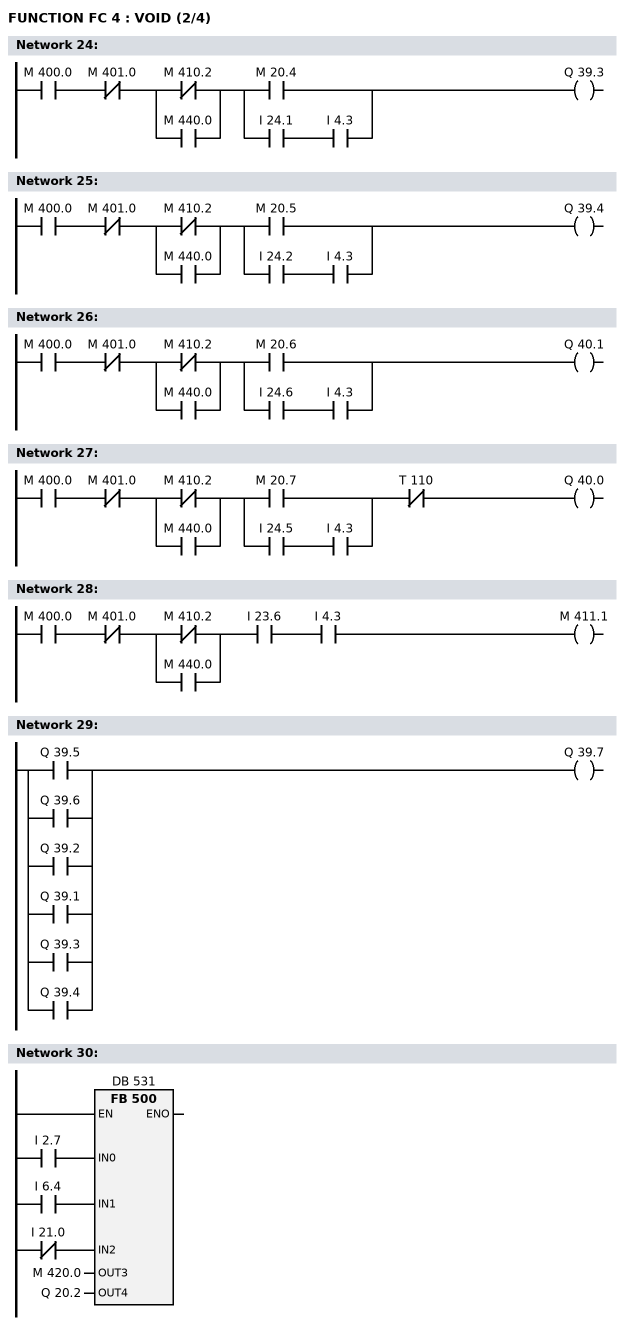

      A     M    400.0;
      AN    M    401.0;
      A(    ;
      ON    M    410.2;
      O     M    440.0;
      )     ;
      A(    ;
      O     M     20.4;
      O     ;
      A     I     24.1;
      A     I      4.3;
      )     ;
      =     Q     39.3;
NETWORK
TITLE =

      A     M    400.0;
      AN    M    401.0;
      A(    ;
      ON    M    410.2;
      O     M    440.0;
      )     ;
      A(    ;
      O     M     20.5;
      O     ;
      A     I     24.2;
      A     I      4.3;
      )     ;
      =     Q     39.4;
NETWORK
TITLE =

      A     M    400.0;
      AN    M    401.0;
      A(    ;
      ON    M    410.2;
      O     M    440.0;
      )     ;
      A(    ;
      O     M     20.6;
      O     ;
      A     I     24.6;
      A     I      4.3;
      )     ;
      =     Q     40.1;
NETWORK
TITLE =

      A     M    400.0;
      AN    M    401.0;
      A(    ;
      ON    M    410.2;
      O     M    440.0;
      )     ;
      A(    ;
      O     M     20.7;
      O     ;
      A     I     24.5;
      A     I      4.3;
      )     ;
      AN    T    110;
      =     Q     40.0;
NETWORK
TITLE =

      A     M    400.0;
      AN    M    401.0;
      A(    ;
      ON    M    410.2;
      O     M    440.0;
      )     ;
      A     I     23.6;
      A     I      4.3;
      =     M    411.1;
NETWORK
TITLE =

      O     Q     39.5;
      O     Q     39.6;
      O     Q     39.2;
      O     Q     39.1;
      O     Q     39.3;
      O     Q     39.4;
      =     Q     39.7;
NETWORK
TITLE =

      A     I      2.7;
      =     L      0.0;
      BLD   103;
      A     I      6.4;
      =     L      0.1;
      BLD   103;
      AN    I     21.0;
      =     L      0.2;
      BLD   103;
      CALL FB   500 , DB   531 (
           IN0                      := L      0.0,
           IN1                      := L      0.1,
           IN2                      := L      0.2,
           OUT3                     := M    420.0,
           OUT4                     := Q     20.2);
      NOP   0;
NETWORK
TITLE =
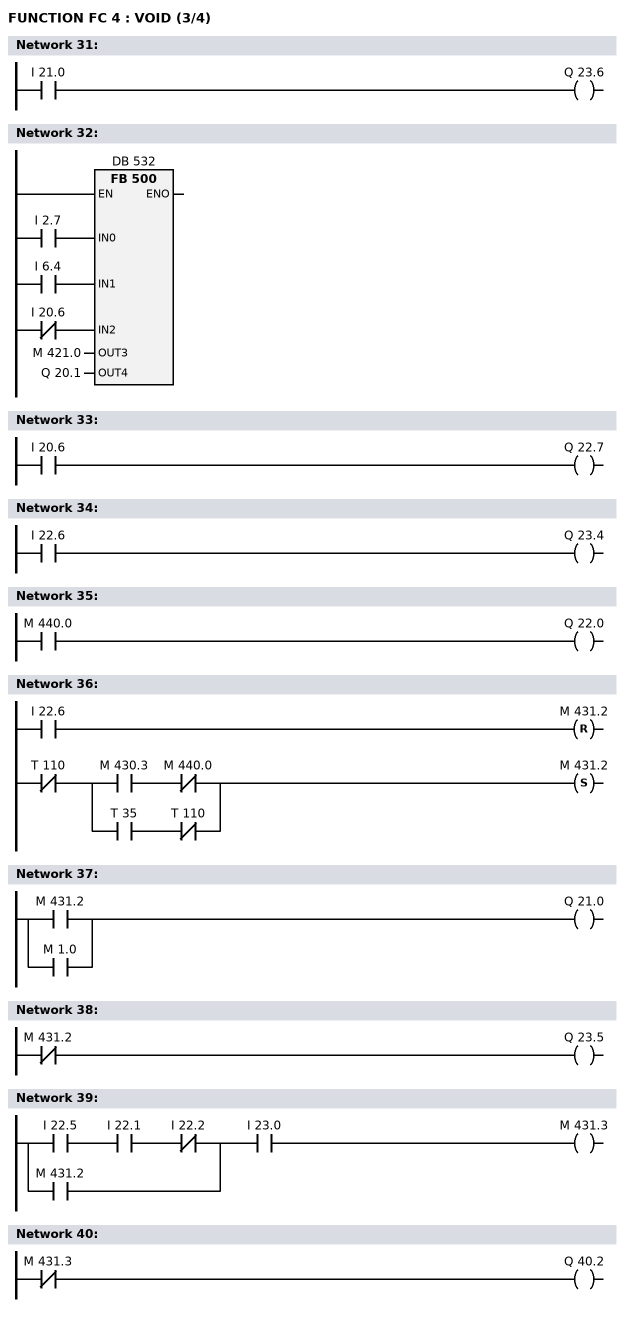

      A     I     21.0;
      =     Q     23.6;
NETWORK
TITLE =

      A     I      2.7;
      =     L      0.0;
      BLD   103;
      A     I      6.4;
      =     L      0.1;
      BLD   103;
      AN    I     20.6;
      =     L      0.2;
      BLD   103;
      CALL FB   500 , DB   532 (
           IN0                      := L      0.0,
           IN1                      := L      0.1,
           IN2                      := L      0.2,
           OUT3                     := M    421.0,
           OUT4                     := Q     20.1);
      NOP   0;
NETWORK
TITLE =

      A     I     20.6;
      =     Q     22.7;
NETWORK
TITLE =

      A     I     22.6;
      =     Q     23.4;
NETWORK
TITLE =

      A     M    440.0;
      =     Q     22.0;
NETWORK
TITLE =

      A     I     22.6;
      R     M    431.2;
      AN    T    110;
      A(    ;
      A     M    430.3;
      AN    M    440.0;
      O     ;
      A     T     35;
      AN    T    110;
      )     ;
      S     M    431.2;
      NOP   0;
NETWORK
TITLE =

      O     M    431.2;
      O     M      1.0;
      =     Q     21.0;
NETWORK
TITLE =

      AN    M    431.2;
      =     Q     23.5;
NETWORK
TITLE =

      A(    ;
      A     I     22.5;
      A     I     22.1;
      AN    I     22.2;
      O     M    431.2;
      )     ;
      A     I     23.0;
      =     M    431.3;
NETWORK
TITLE =

      AN    M    431.3;
      =     Q     40.2;
NETWORK
TITLE =
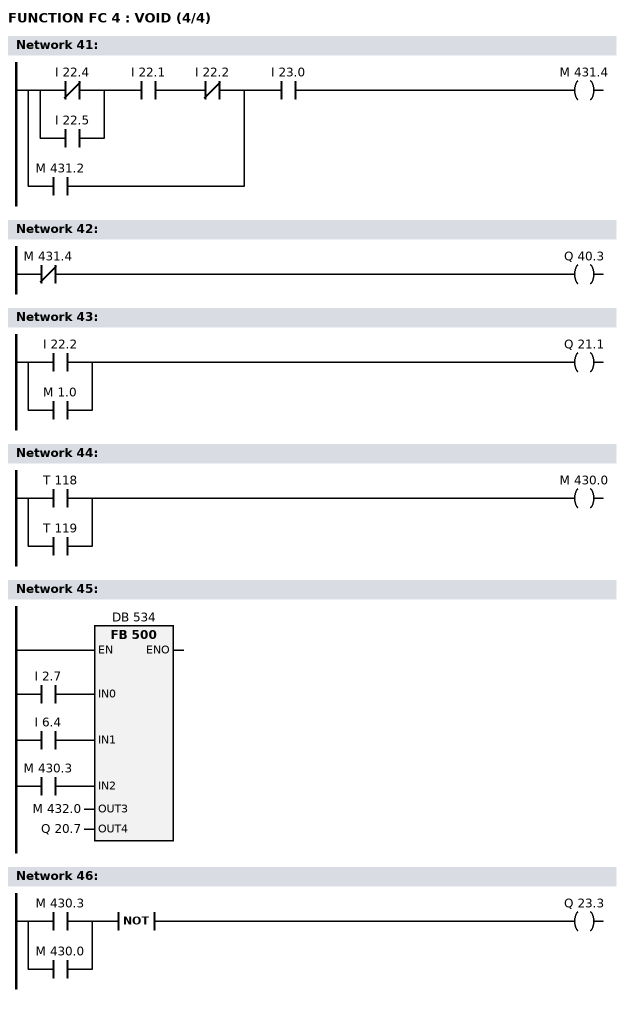

      A(    ;
      A(    ;
      ON    I     22.4;
      O     I     22.5;
      )     ;
      A     I     22.1;
      AN    I     22.2;
      O     M    431.2;
      )     ;
      A     I     23.0;
      =     M    431.4;
NETWORK
TITLE =

      AN    M    431.4;
      =     Q     40.3;
NETWORK
TITLE =

      O     I     22.2;
      O     M      1.0;
      =     Q     21.1;
NETWORK
TITLE =

      O     T    118;
      O     T    119;
      =     M    430.0;
NETWORK
TITLE =

      A     I      2.7;
      =     L      0.0;
      BLD   103;
      A     I      6.4;
      =     L      0.1;
      BLD   103;
      A     M    430.3;
      =     L      0.2;
      BLD   103;
      CALL FB   500 , DB   534 (
           IN0                      := L      0.0,
           IN1                      := L      0.1,
           IN2                      := L      0.2,
           OUT3                     := M    432.0,
           OUT4                     := Q     20.7);
      NOP   0;
NETWORK
TITLE =

      A(    ;
      O     M    430.3;
      O     M    430.0;
      )     ;
      NOT   ;
      =     Q     23.3;
NETWORK
TITLE =

      A(    ;
      A     I     21.5;
      L     S5T#150MS;
      SD    T    103;
      NOP   0;
      NOP   0;
      NOP   0;
      A     T    103;
      )     ;
      NOT   ;
      =     Q     21.6;
NETWORK
TITLE =

      A(    ;
      A     I     21.7;
      L     S5T#150MS;
      SD    T    104;
      NOP   0;
      NOP   0;
      NOP   0;
      A     T    104;
      )     ;
      NOT   ;
      =     Q     23.1;
NETWORK
TITLE =

      A(    ;
      A     I     21.6;
      L     S5T#150MS;
      SD    T    106;
      NOP   0;
      NOP   0;
      NOP   0;
      A     T    106;
      )     ;
      NOT   ;
      =     Q     22.6;
NETWORK
TITLE =

      A(    ;
      A     I     21.4;
      L     S5T#150MS;
      SD    T    107;
      NOP   0;
      NOP   0;
      NOP   0;
      A     T    107;
      )     ;
      NOT   ;
      =     Q     23.2;
NETWORK
TITLE =
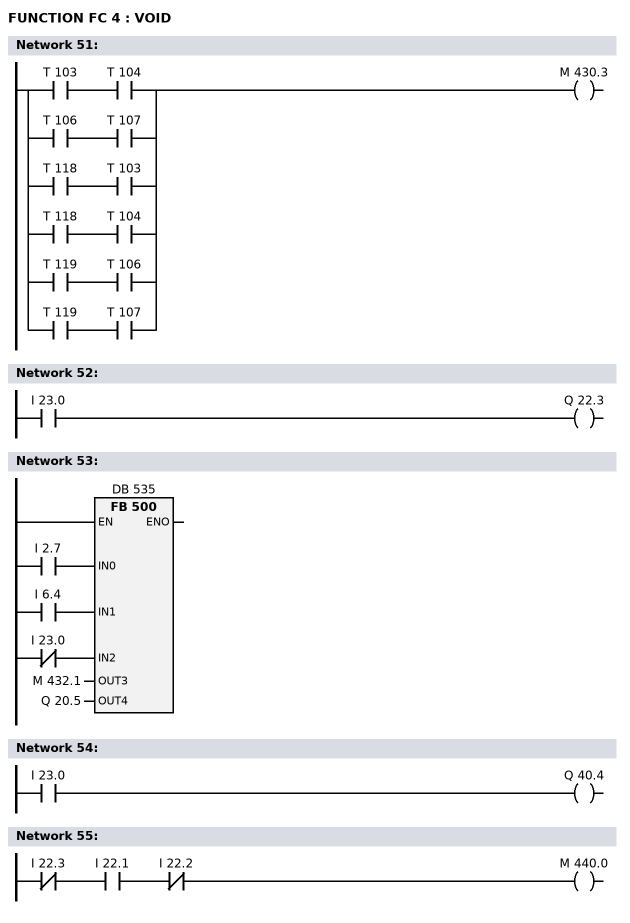

      A     T    103;
      A     T    104;
      O     ;
      A     T    106;
      A     T    107;
      O     ;
      A     T    118;
      A     T    103;
      O     ;
      A     T    118;
      A     T    104;
      O     ;
      A     T    119;
      A     T    106;
      O     ;
      A     T    119;
      A     T    107;
      =     M    430.3;
NETWORK
TITLE =

      A     I     23.0;
      =     Q     22.3;
NETWORK
TITLE =

      A     I      2.7;
      =     L      0.0;
      BLD   103;
      A     I      6.4;
      =     L      0.1;
      BLD   103;
      AN    I     23.0;
      =     L      0.2;
      BLD   103;
      CALL FB   500 , DB   535 (
           IN0                      := L      0.0,
           IN1                      := L      0.1,
           IN2                      := L      0.2,
           OUT3                     := M    432.1,
           OUT4                     := Q     20.5);
      NOP   0;
NETWORK
TITLE =

      A     I     23.0;
      =     Q     40.4;
NETWORK
TITLE =

      AN    I     22.3;
      A     I     22.1;
      AN    I     22.2;
      =     M    440.0;
END_FUNCTION

FUNCTION FC 5 : VOID
VERSION : 0.1

BEGIN
NETWORK
TITLE =
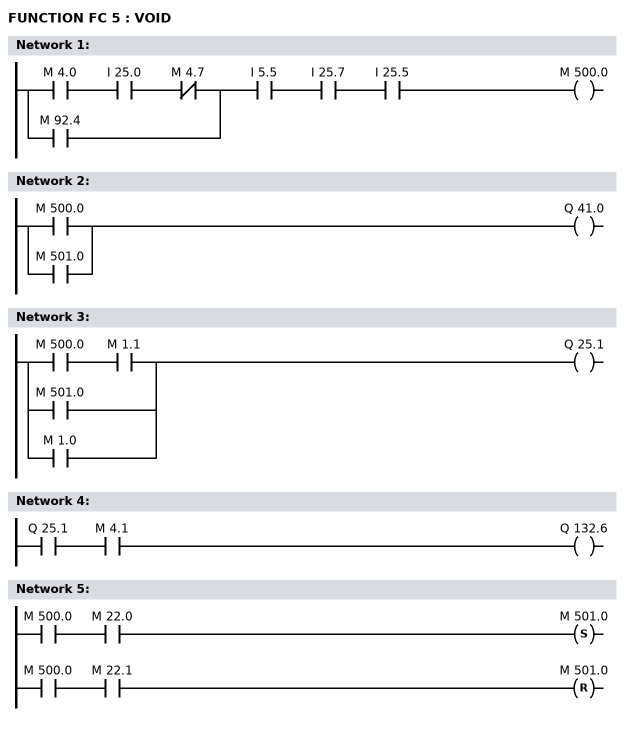

      A(    ;
      A     M      4.0;
      A     I     25.0;
      AN    M      4.7;
      O     M     92.4;
      )     ;
      A     I      5.5;
      A     I     25.7;
      A     I     25.5;
      =     M    500.0;
NETWORK
TITLE =

      O     M    500.0;
      O     M    501.0;
      =     Q     41.0;
NETWORK
TITLE =

      A     M    500.0;
      A     M      1.1;
      O     M    501.0;
      O     M      1.0;
      =     Q     25.1;
NETWORK
TITLE =

      A     Q     25.1;
      A     M      4.1;
      =     Q    132.6;
NETWORK
TITLE =

      A     M    500.0;
      A     M     22.0;
      S     M    501.0;
      A     M    500.0;
      A     M     22.1;
      R     M    501.0;
      NOP   0;
NETWORK
TITLE =

      A(    ;
      A     I     25.3;
      L     S5T#150MS;
      SD    T    128;
      NOP   0;
      NOP   0;
      NOP   0;
      A     T    128;
      )     ;
      NOT   ;
      =     Q     25.7;
NETWORK
TITLE =

      A(    ;
      A     I     25.2;
      L     S5T#150MS;
      SD    T    129;
      NOP   0;
      NOP   0;
      NOP   0;
      A     T    129;
      )     ;
      NOT   ;
      =     Q     25.6;
NETWORK
TITLE =
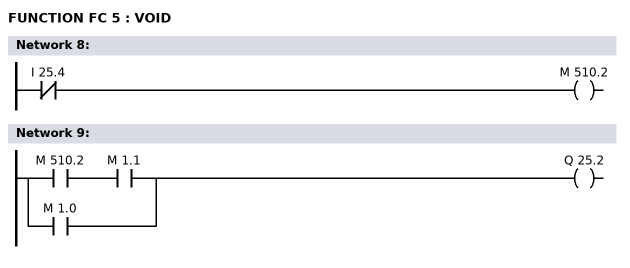

      AN    I     25.4;
      =     M    510.2;
NETWORK
TITLE =

      A     M    510.2;
      A     M      1.1;
      O     M      1.0;
      =     Q     25.2;
NETWORK
TITLE =

      O(    ;
      A     I     25.1;
      L     S5T#150MS;
      SD    T    130;
      NOP   0;
      NOP   0;
      NOP   0;
      A     T    130;
      )     ;
      O     M      1.0;
      =     Q     25.0;
NETWORK
TITLE =
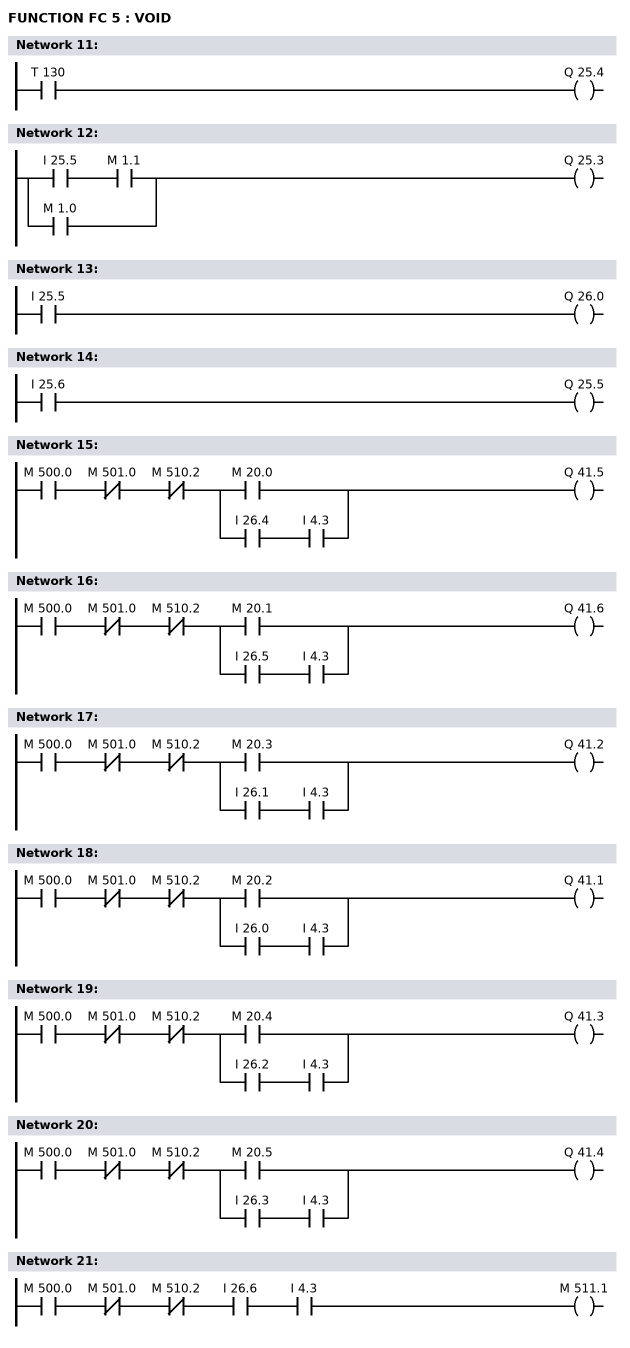

      A     T    130;
      =     Q     25.4;
NETWORK
TITLE =

      A     I     25.5;
      A     M      1.1;
      O     M      1.0;
      =     Q     25.3;
NETWORK
TITLE =

      A     I     25.5;
      =     Q     26.0;
NETWORK
TITLE =

      A     I     25.6;
      =     Q     25.5;
NETWORK
TITLE =

      A     M    500.0;
      AN    M    501.0;
      AN    M    510.2;
      A(    ;
      O     M     20.0;
      O     ;
      A     I     26.4;
      A     I      4.3;
      )     ;
      =     Q     41.5;
NETWORK
TITLE =

      A     M    500.0;
      AN    M    501.0;
      AN    M    510.2;
      A(    ;
      O     M     20.1;
      O     ;
      A     I     26.5;
      A     I      4.3;
      )     ;
      =     Q     41.6;
NETWORK
TITLE =

      A     M    500.0;
      AN    M    501.0;
      AN    M    510.2;
      A(    ;
      O     M     20.3;
      O     ;
      A     I     26.1;
      A     I      4.3;
      )     ;
      =     Q     41.2;
NETWORK
TITLE =

      A     M    500.0;
      AN    M    501.0;
      AN    M    510.2;
      A(    ;
      O     M     20.2;
      O     ;
      A     I     26.0;
      A     I      4.3;
      )     ;
      =     Q     41.1;
NETWORK
TITLE =

      A     M    500.0;
      AN    M    501.0;
      AN    M    510.2;
      A(    ;
      O     M     20.4;
      O     ;
      A     I     26.2;
      A     I      4.3;
      )     ;
      =     Q     41.3;
NETWORK
TITLE =

      A     M    500.0;
      AN    M    501.0;
      AN    M    510.2;
      A(    ;
      O     M     20.5;
      O     ;
      A     I     26.3;
      A     I      4.3;
      )     ;
      =     Q     41.4;
NETWORK
TITLE =

      A     M    500.0;
      AN    M    501.0;
      AN    M    510.2;
      A     I     26.6;
      A     I      4.3;
      =     M    511.1;
END_FUNCTION

FUNCTION FC 6 : VOID
VERSION : 0.1

BEGIN
NETWORK
TITLE =
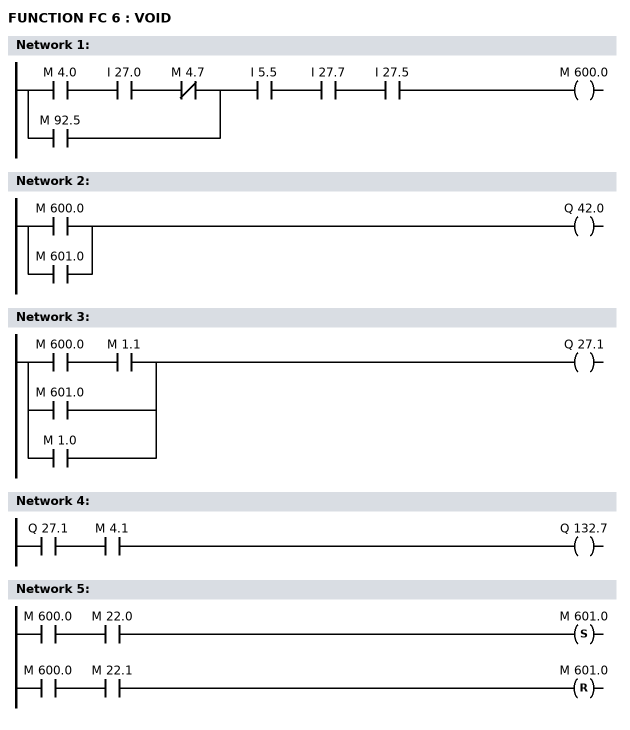

      A(    ;
      A     M      4.0;
      A     I     27.0;
      AN    M      4.7;
      O     M     92.5;
      )     ;
      A     I      5.5;
      A     I     27.7;
      A     I     27.5;
      =     M    600.0;
NETWORK
TITLE =

      O     M    600.0;
      O     M    601.0;
      =     Q     42.0;
NETWORK
TITLE =

      A     M    600.0;
      A     M      1.1;
      O     M    601.0;
      O     M      1.0;
      =     Q     27.1;
NETWORK
TITLE =

      A     Q     27.1;
      A     M      4.1;
      =     Q    132.7;
NETWORK
TITLE =

      A     M    600.0;
      A     M     22.0;
      S     M    601.0;
      A     M    600.0;
      A     M     22.1;
      R     M    601.0;
      NOP   0;
NETWORK
TITLE =

      A(    ;
      A     I     27.3;
      L     S5T#150MS;
      SD    T    148;
      NOP   0;
      NOP   0;
      NOP   0;
      A     T    148;
      )     ;
      NOT   ;
      =     Q     27.7;
NETWORK
TITLE =

      A(    ;
      A     I     27.2;
      L     S5T#150MS;
      SD    T    149;
      NOP   0;
      NOP   0;
      NOP   0;
      A     T    149;
      )     ;
      NOT   ;
      =     Q     27.6;
NETWORK
TITLE =
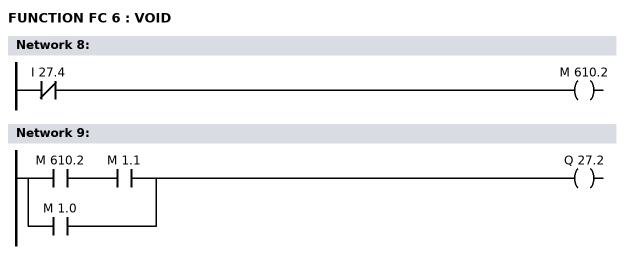

      AN    I     27.4;
      =     M    610.2;
NETWORK
TITLE =

      A     M    610.2;
      A     M      1.1;
      O     M      1.0;
      =     Q     27.2;
NETWORK
TITLE =

      O(    ;
      A     I     27.1;
      L     S5T#150MS;
      SD    T    150;
      NOP   0;
      NOP   0;
      NOP   0;
      A     T    150;
      )     ;
      O     M      1.0;
      =     Q     27.0;
NETWORK
TITLE =
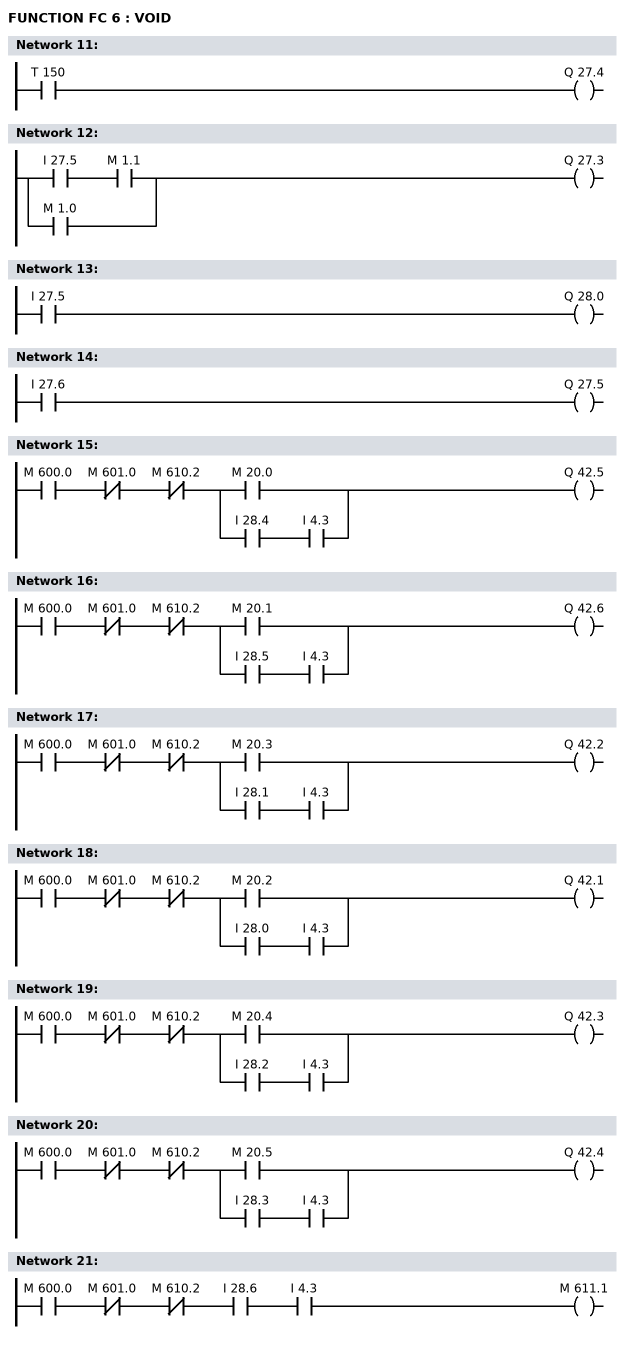

      A     T    150;
      =     Q     27.4;
NETWORK
TITLE =

      A     I     27.5;
      A     M      1.1;
      O     M      1.0;
      =     Q     27.3;
NETWORK
TITLE =

      A     I     27.5;
      =     Q     28.0;
NETWORK
TITLE =

      A     I     27.6;
      =     Q     27.5;
NETWORK
TITLE =

      A     M    600.0;
      AN    M    601.0;
      AN    M    610.2;
      A(    ;
      O     M     20.0;
      O     ;
      A     I     28.4;
      A     I      4.3;
      )     ;
      =     Q     42.5;
NETWORK
TITLE =

      A     M    600.0;
      AN    M    601.0;
      AN    M    610.2;
      A(    ;
      O     M     20.1;
      O     ;
      A     I     28.5;
      A     I      4.3;
      )     ;
      =     Q     42.6;
NETWORK
TITLE =

      A     M    600.0;
      AN    M    601.0;
      AN    M    610.2;
      A(    ;
      O     M     20.3;
      O     ;
      A     I     28.1;
      A     I      4.3;
      )     ;
      =     Q     42.2;
NETWORK
TITLE =

      A     M    600.0;
      AN    M    601.0;
      AN    M    610.2;
      A(    ;
      O     M     20.2;
      O     ;
      A     I     28.0;
      A     I      4.3;
      )     ;
      =     Q     42.1;
NETWORK
TITLE =

      A     M    600.0;
      AN    M    601.0;
      AN    M    610.2;
      A(    ;
      O     M     20.4;
      O     ;
      A     I     28.2;
      A     I      4.3;
      )     ;
      =     Q     42.3;
NETWORK
TITLE =

      A     M    600.0;
      AN    M    601.0;
      AN    M    610.2;
      A(    ;
      O     M     20.5;
      O     ;
      A     I     28.3;
      A     I      4.3;
      )     ;
      =     Q     42.4;
NETWORK
TITLE =

      A     M    600.0;
      AN    M    601.0;
      AN    M    610.2;
      A     I     28.6;
      A     I      4.3;
      =     M    611.1;
END_FUNCTION

FUNCTION FC 7 : VOID
VERSION : 0.1

BEGIN
NETWORK
TITLE =
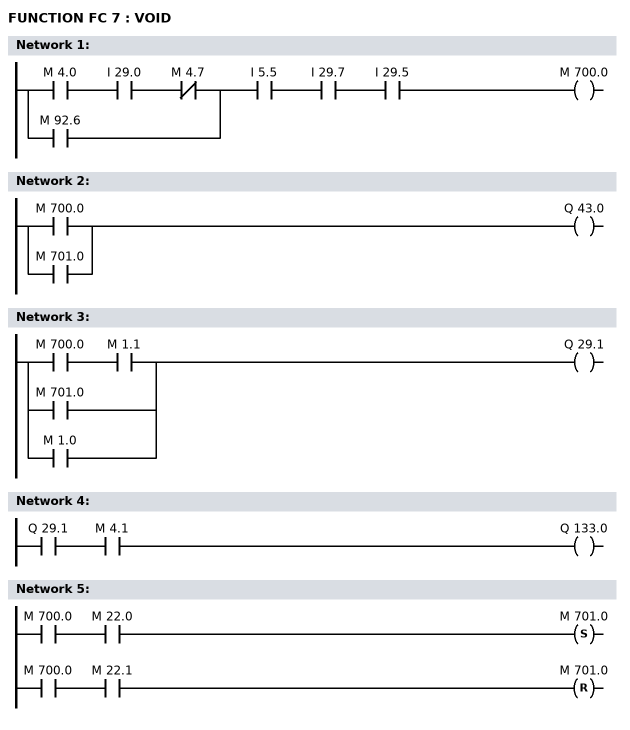

      A(    ;
      A     M      4.0;
      A     I     29.0;
      AN    M      4.7;
      O     M     92.6;
      )     ;
      A     I      5.5;
      A     I     29.7;
      A     I     29.5;
      =     M    700.0;
NETWORK
TITLE =

      O     M    700.0;
      O     M    701.0;
      =     Q     43.0;
NETWORK
TITLE =

      A     M    700.0;
      A     M      1.1;
      O     M    701.0;
      O     M      1.0;
      =     Q     29.1;
NETWORK
TITLE =

      A     Q     29.1;
      A     M      4.1;
      =     Q    133.0;
NETWORK
TITLE =

      A     M    700.0;
      A     M     22.0;
      S     M    701.0;
      A     M    700.0;
      A     M     22.1;
      R     M    701.0;
      NOP   0;
NETWORK
TITLE =

      A(    ;
      A     I     29.3;
      L     S5T#150MS;
      SD    T    168;
      NOP   0;
      NOP   0;
      NOP   0;
      A     T    168;
      )     ;
      NOT   ;
      =     Q     29.7;
NETWORK
TITLE =

      A(    ;
      A     I     29.2;
      L     S5T#150MS;
      SD    T    169;
      NOP   0;
      NOP   0;
      NOP   0;
      A     T    169;
      )     ;
      NOT   ;
      =     Q     29.6;
NETWORK
TITLE =
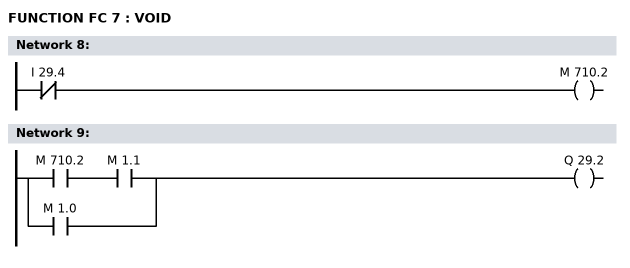

      AN    I     29.4;
      =     M    710.2;
NETWORK
TITLE =

      A     M    710.2;
      A     M      1.1;
      O     M      1.0;
      =     Q     29.2;
NETWORK
TITLE =

      O(    ;
      A     I     29.1;
      L     S5T#150MS;
      SD    T    170;
      NOP   0;
      NOP   0;
      NOP   0;
      A     T    170;
      )     ;
      O     M      1.0;
      =     Q     29.0;
NETWORK
TITLE =
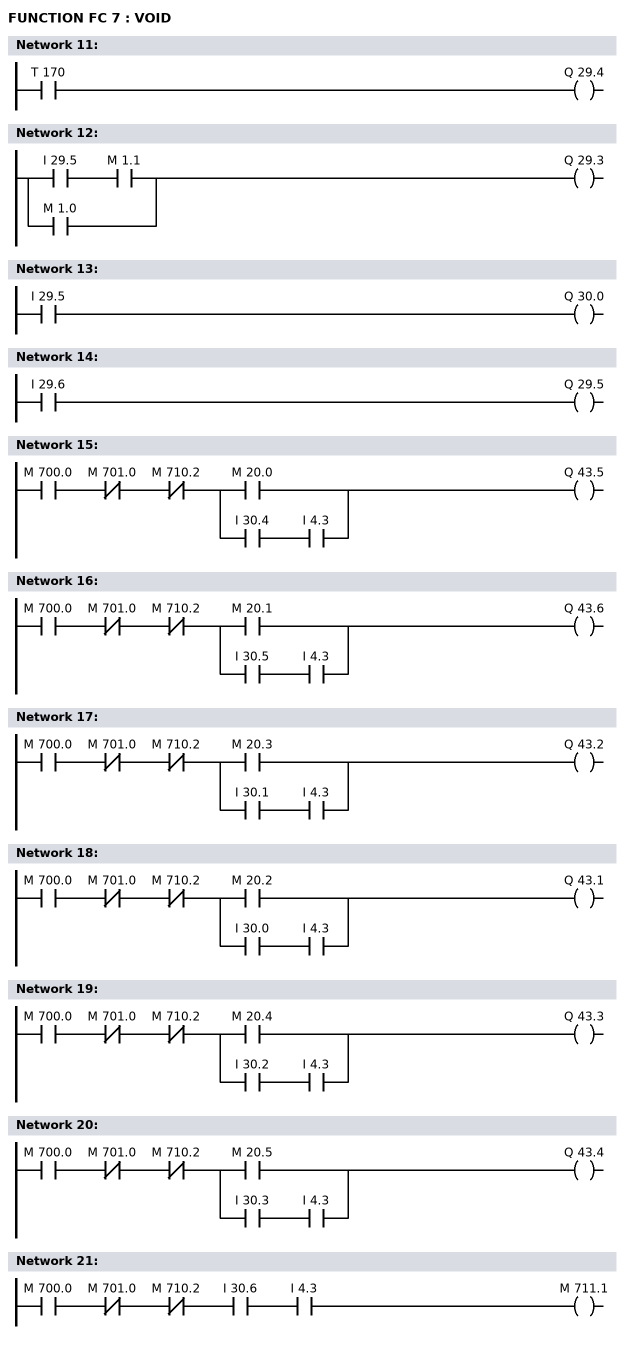

      A     T    170;
      =     Q     29.4;
NETWORK
TITLE =

      A     I     29.5;
      A     M      1.1;
      O     M      1.0;
      =     Q     29.3;
NETWORK
TITLE =

      A     I     29.5;
      =     Q     30.0;
NETWORK
TITLE =

      A     I     29.6;
      =     Q     29.5;
NETWORK
TITLE =

      A     M    700.0;
      AN    M    701.0;
      AN    M    710.2;
      A(    ;
      O     M     20.0;
      O     ;
      A     I     30.4;
      A     I      4.3;
      )     ;
      =     Q     43.5;
NETWORK
TITLE =

      A     M    700.0;
      AN    M    701.0;
      AN    M    710.2;
      A(    ;
      O     M     20.1;
      O     ;
      A     I     30.5;
      A     I      4.3;
      )     ;
      =     Q     43.6;
NETWORK
TITLE =

      A     M    700.0;
      AN    M    701.0;
      AN    M    710.2;
      A(    ;
      O     M     20.3;
      O     ;
      A     I     30.1;
      A     I      4.3;
      )     ;
      =     Q     43.2;
NETWORK
TITLE =

      A     M    700.0;
      AN    M    701.0;
      AN    M    710.2;
      A(    ;
      O     M     20.2;
      O     ;
      A     I     30.0;
      A     I      4.3;
      )     ;
      =     Q     43.1;
NETWORK
TITLE =

      A     M    700.0;
      AN    M    701.0;
      AN    M    710.2;
      A(    ;
      O     M     20.4;
      O     ;
      A     I     30.2;
      A     I      4.3;
      )     ;
      =     Q     43.3;
NETWORK
TITLE =

      A     M    700.0;
      AN    M    701.0;
      AN    M    710.2;
      A(    ;
      O     M     20.5;
      O     ;
      A     I     30.3;
      A     I      4.3;
      )     ;
      =     Q     43.4;
NETWORK
TITLE =

      A     M    700.0;
      AN    M    701.0;
      AN    M    710.2;
      A     I     30.6;
      A     I      4.3;
      =     M    711.1;
END_FUNCTION

FUNCTION FC 11 : VOID
VERSION : 0.1

BEGIN
NETWORK
TITLE =
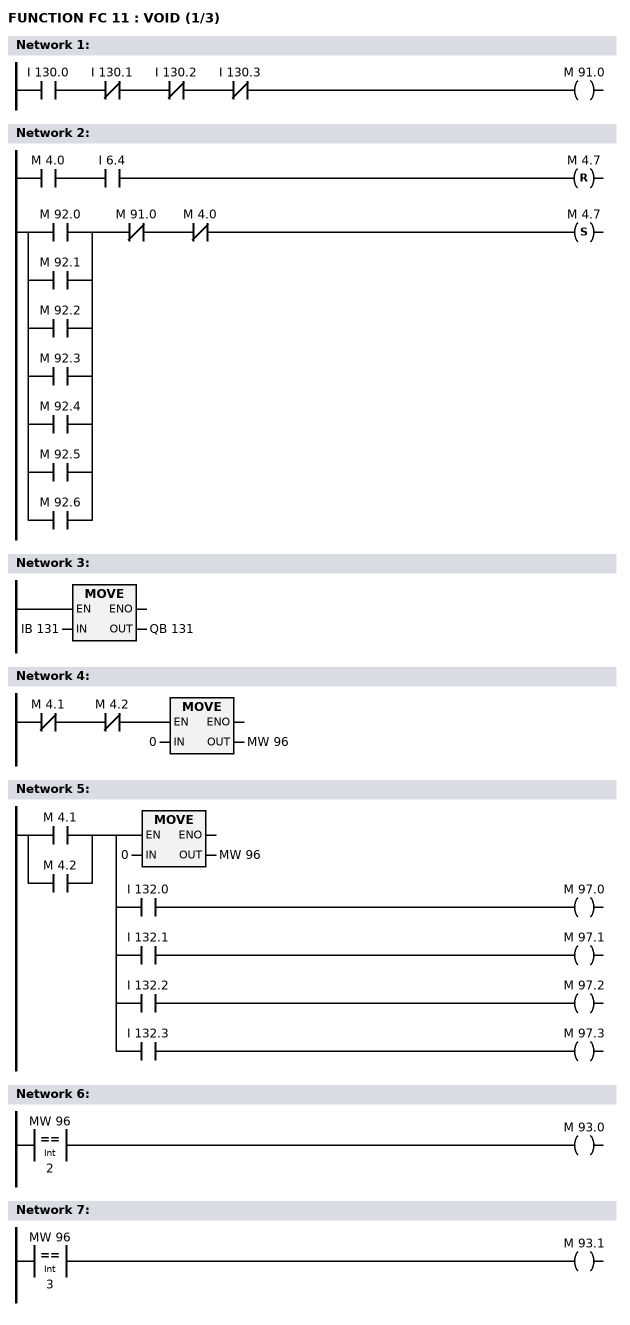

      A     I    130.0;
      AN    I    130.1;
      AN    I    130.2;
      AN    I    130.3;
      =     M     91.0;
NETWORK
TITLE =

      A     M      4.0;
      A     I      6.4;
      R     M      4.7;
      A(    ;
      O     M     92.0;
      O     M     92.1;
      O     M     92.2;
      O     M     92.3;
      O     M     92.4;
      O     M     92.5;
      O     M     92.6;
      )     ;
      AN    M     91.0;
      AN    M      4.0;
      S     M      4.7;
      NOP   0;
NETWORK
TITLE =

      L     IB   131;
      T     QB   131;
      NOP   0;
NETWORK
TITLE =

      AN    M      4.1;
      AN    M      4.2;
      JNB   M001;
      L     0;
      T     MW    96;
M001: NOP   0;
NETWORK
TITLE =

      O     M      4.1;
      O     M      4.2;
      =     L      0.0;
      A     L      0.0;
      JNB   M002;
      L     0;
      T     MW    96;
M002: NOP   0;
      A     L      0.0;
      A     I    132.0;
      =     M     97.0;
      A     L      0.0;
      A     I    132.1;
      =     M     97.1;
      A     L      0.0;
      A     I    132.2;
      =     M     97.2;
      A     L      0.0;
      A     I    132.3;
      =     M     97.3;
NETWORK
TITLE =

      L     MW    96;
      L     2;
      ==I   ;
      =     M     93.0;
NETWORK
TITLE =

      L     MW    96;
      L     3;
      ==I   ;
      =     M     93.1;
NETWORK
TITLE =
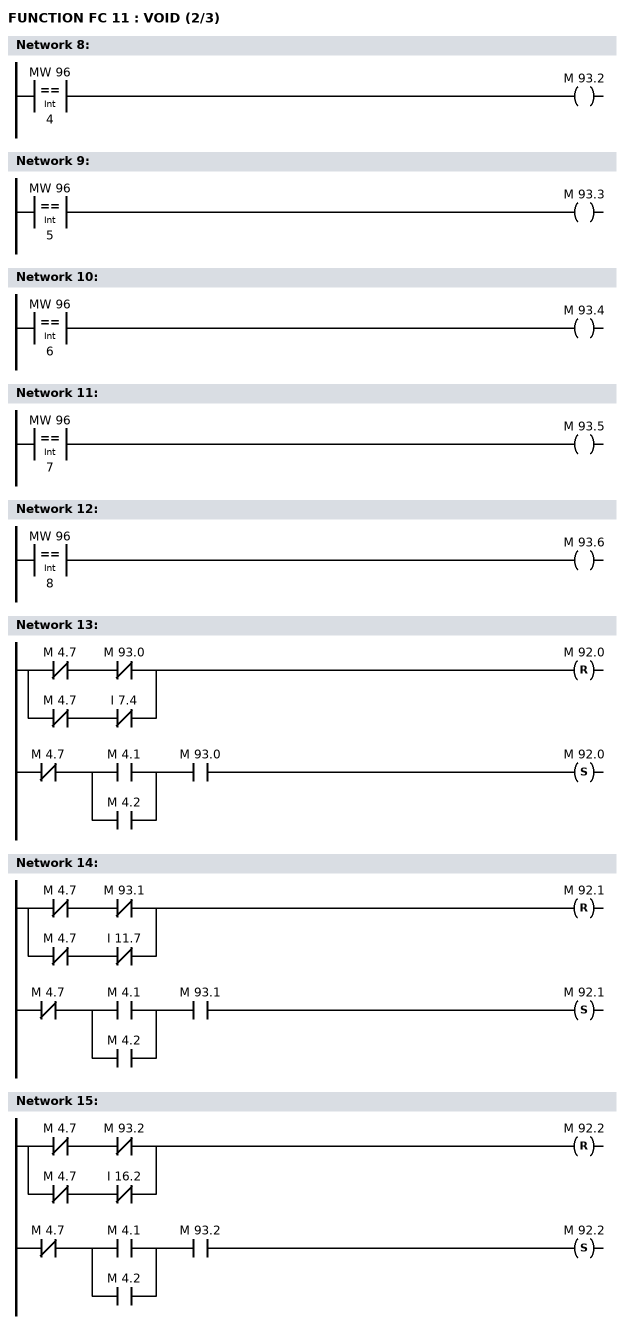

      L     MW    96;
      L     4;
      ==I   ;
      =     M     93.2;
NETWORK
TITLE =

      L     MW    96;
      L     5;
      ==I   ;
      =     M     93.3;
NETWORK
TITLE =

      L     MW    96;
      L     6;
      ==I   ;
      =     M     93.4;
NETWORK
TITLE =

      L     MW    96;
      L     7;
      ==I   ;
      =     M     93.5;
NETWORK
TITLE =

      L     MW    96;
      L     8;
      ==I   ;
      =     M     93.6;
NETWORK
TITLE =

      A(    ;
      AN    M      4.7;
      AN    M     93.0;
      O     ;
      AN    M      4.7;
      AN    I      7.4;
      )     ;
      R     M     92.0;
      AN    M      4.7;
      A(    ;
      O     M      4.1;
      O     M      4.2;
      )     ;
      A     M     93.0;
      S     M     92.0;
      NOP   0;
NETWORK
TITLE =

      A(    ;
      AN    M      4.7;
      AN    M     93.1;
      O     ;
      AN    M      4.7;
      AN    I     11.7;
      )     ;
      R     M     92.1;
      AN    M      4.7;
      A(    ;
      O     M      4.1;
      O     M      4.2;
      )     ;
      A     M     93.1;
      S     M     92.1;
      NOP   0;
NETWORK
TITLE =

      A(    ;
      AN    M      4.7;
      AN    M     93.2;
      O     ;
      AN    M      4.7;
      AN    I     16.2;
      )     ;
      R     M     92.2;
      AN    M      4.7;
      A(    ;
      O     M      4.1;
      O     M      4.2;
      )     ;
      A     M     93.2;
      S     M     92.2;
      NOP   0;
NETWORK
TITLE =
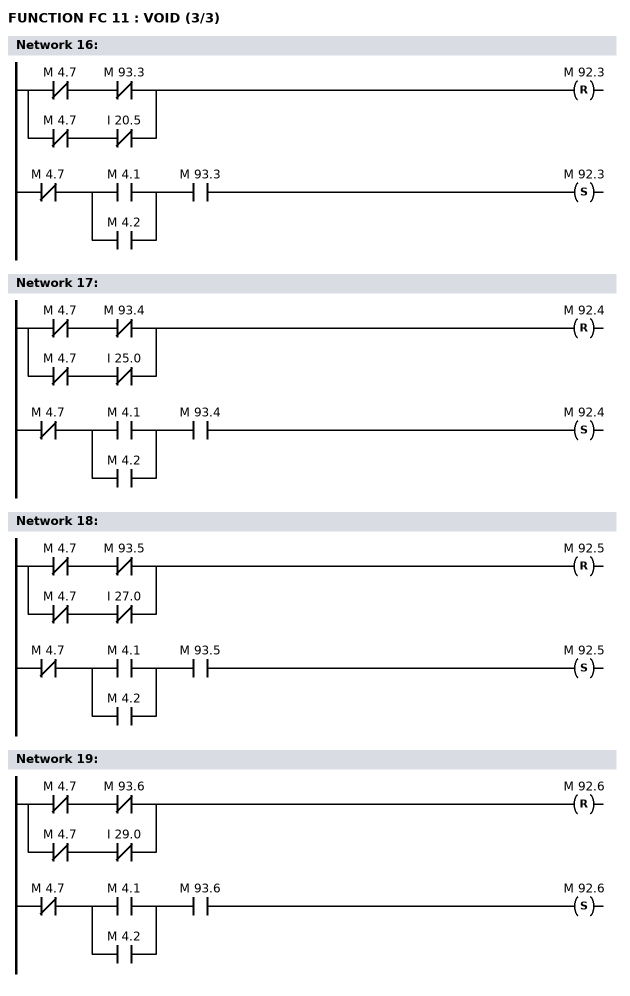

      A(    ;
      AN    M      4.7;
      AN    M     93.3;
      O     ;
      AN    M      4.7;
      AN    I     20.5;
      )     ;
      R     M     92.3;
      AN    M      4.7;
      A(    ;
      O     M      4.1;
      O     M      4.2;
      )     ;
      A     M     93.3;
      S     M     92.3;
      NOP   0;
NETWORK
TITLE =

      A(    ;
      AN    M      4.7;
      AN    M     93.4;
      O     ;
      AN    M      4.7;
      AN    I     25.0;
      )     ;
      R     M     92.4;
      AN    M      4.7;
      A(    ;
      O     M      4.1;
      O     M      4.2;
      )     ;
      A     M     93.4;
      S     M     92.4;
      NOP   0;
NETWORK
TITLE =

      A(    ;
      AN    M      4.7;
      AN    M     93.5;
      O     ;
      AN    M      4.7;
      AN    I     27.0;
      )     ;
      R     M     92.5;
      AN    M      4.7;
      A(    ;
      O     M      4.1;
      O     M      4.2;
      )     ;
      A     M     93.5;
      S     M     92.5;
      NOP   0;
NETWORK
TITLE =

      A(    ;
      AN    M      4.7;
      AN    M     93.6;
      O     ;
      AN    M      4.7;
      AN    I     29.0;
      )     ;
      R     M     92.6;
      AN    M      4.7;
      A(    ;
      O     M      4.1;
      O     M      4.2;
      )     ;
      A     M     93.6;
      S     M     92.6;
      NOP   0;
END_FUNCTION

FUNCTION FC 13 : VOID
VERSION : 0.1

BEGIN
NETWORK
TITLE =
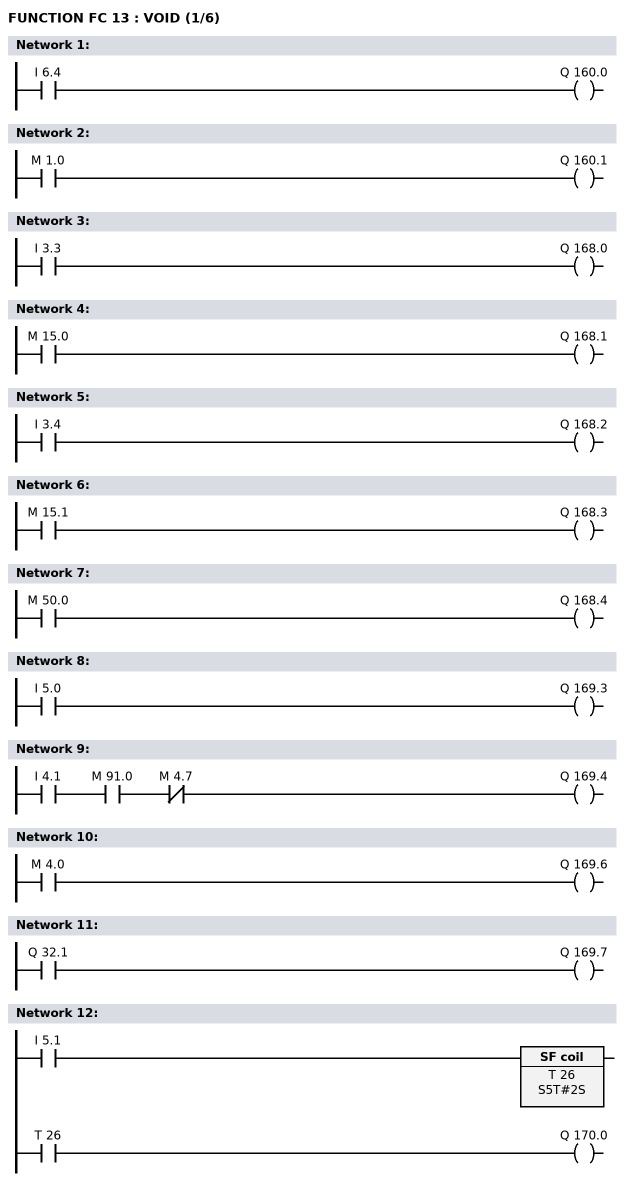

      A     I      6.4;
      =     Q    160.0;
NETWORK
TITLE =

      A     M      1.0;
      =     Q    160.1;
NETWORK
TITLE =

      A     I      3.3;
      =     Q    168.0;
NETWORK
TITLE =

      A     M     15.0;
      =     Q    168.1;
NETWORK
TITLE =

      A     I      3.4;
      =     Q    168.2;
NETWORK
TITLE =

      A     M     15.1;
      =     Q    168.3;
NETWORK
TITLE =

      A     M     50.0;
      =     Q    168.4;
NETWORK
TITLE =

      A     I      5.0;
      =     Q    169.3;
NETWORK
TITLE =

      A     I      4.1;
      A     M     91.0;
      AN    M      4.7;
      =     Q    169.4;
NETWORK
TITLE =

      A     M      4.0;
      =     Q    169.6;
NETWORK
TITLE =

      A     Q     32.1;
      =     Q    169.7;
NETWORK
TITLE =

      A     I      5.1;
      L     S5T#2S;
      SF    T     26;
      NOP   0;
      NOP   0;
      NOP   0;
      A     T     26;
      =     Q    170.0;
NETWORK
TITLE =
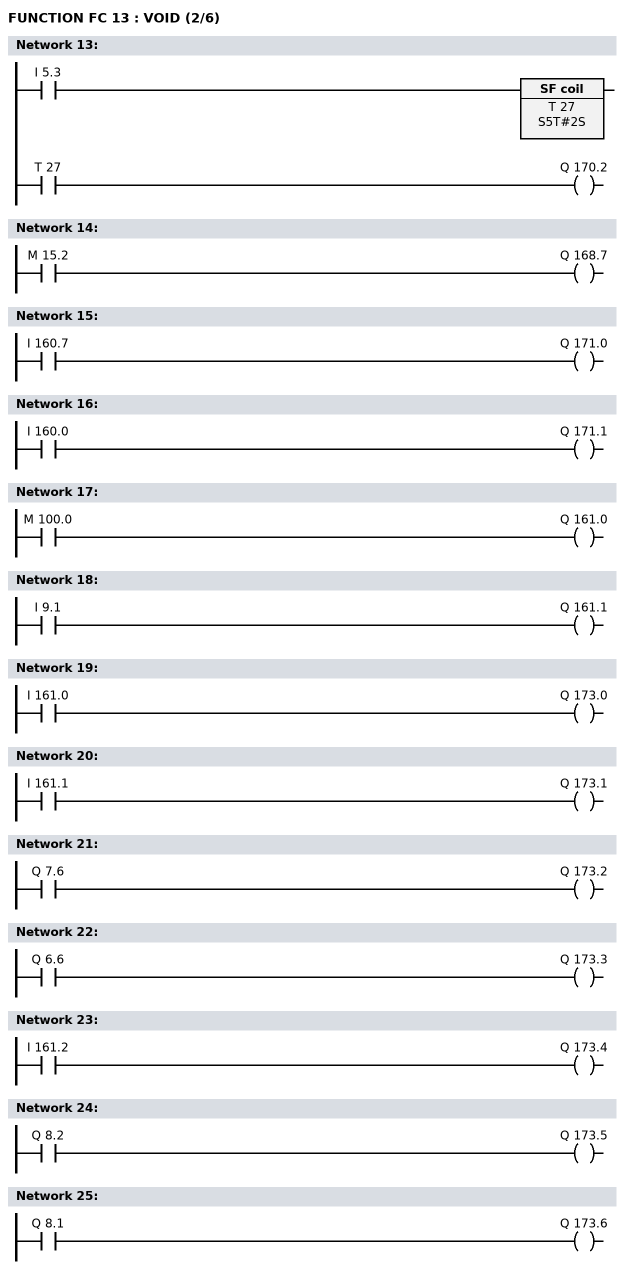

      A     I      5.3;
      L     S5T#2S;
      SF    T     27;
      NOP   0;
      NOP   0;
      NOP   0;
      A     T     27;
      =     Q    170.2;
NETWORK
TITLE =

      A     M     15.2;
      =     Q    168.7;
NETWORK
TITLE =

      A     I    160.7;
      =     Q    171.0;
NETWORK
TITLE =

      A     I    160.0;
      =     Q    171.1;
NETWORK
TITLE =

      A     M    100.0;
      =     Q    161.0;
NETWORK
TITLE =

      A     I      9.1;
      =     Q    161.1;
NETWORK
TITLE =

      A     I    161.0;
      =     Q    173.0;
NETWORK
TITLE =

      A     I    161.1;
      =     Q    173.1;
NETWORK
TITLE =

      A     Q      7.6;
      =     Q    173.2;
NETWORK
TITLE =

      A     Q      6.6;
      =     Q    173.3;
NETWORK
TITLE =

      A     I    161.2;
      =     Q    173.4;
NETWORK
TITLE =

      A     Q      8.2;
      =     Q    173.5;
NETWORK
TITLE =

      A     Q      8.1;
      =     Q    173.6;
NETWORK
TITLE =
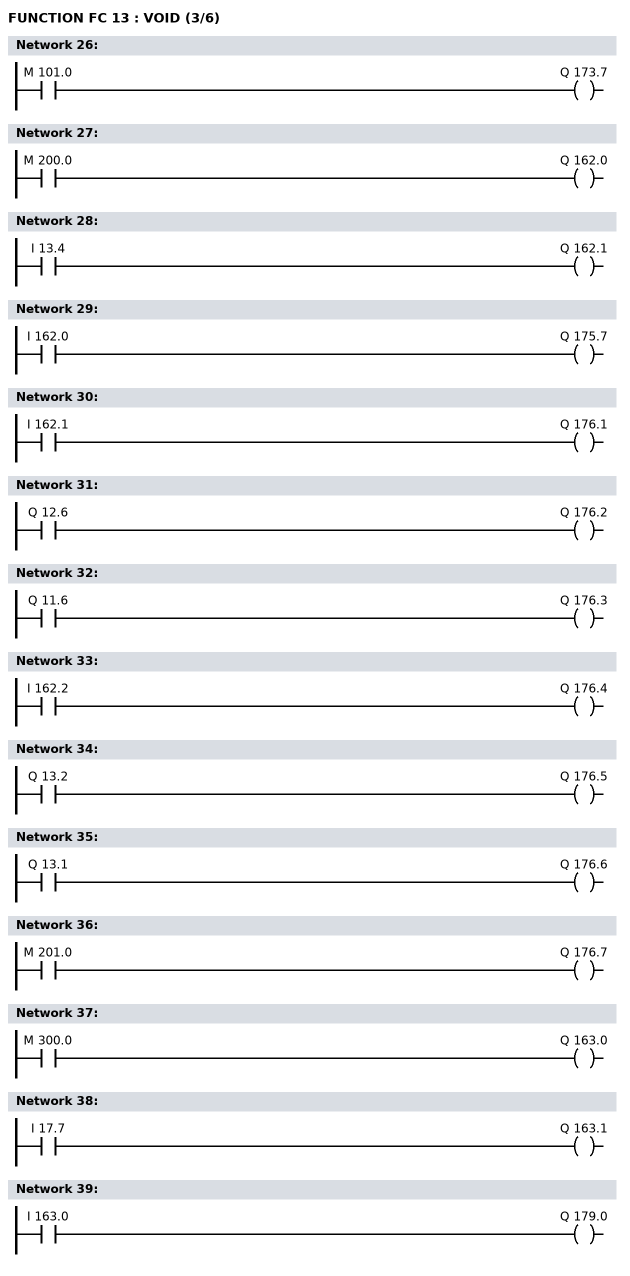

      A     M    101.0;
      =     Q    173.7;
NETWORK
TITLE =

      A     M    200.0;
      =     Q    162.0;
NETWORK
TITLE =

      A     I     13.4;
      =     Q    162.1;
NETWORK
TITLE =

      A     I    162.0;
      =     Q    175.7;
NETWORK
TITLE =

      A     I    162.1;
      =     Q    176.1;
NETWORK
TITLE =

      A     Q     12.6;
      =     Q    176.2;
NETWORK
TITLE =

      A     Q     11.6;
      =     Q    176.3;
NETWORK
TITLE =

      A     I    162.2;
      =     Q    176.4;
NETWORK
TITLE =

      A     Q     13.2;
      =     Q    176.5;
NETWORK
TITLE =

      A     Q     13.1;
      =     Q    176.6;
NETWORK
TITLE =

      A     M    201.0;
      =     Q    176.7;
NETWORK
TITLE =

      A     M    300.0;
      =     Q    163.0;
NETWORK
TITLE =

      A     I     17.7;
      =     Q    163.1;
NETWORK
TITLE =

      A     I    163.0;
      =     Q    179.0;
NETWORK
TITLE =
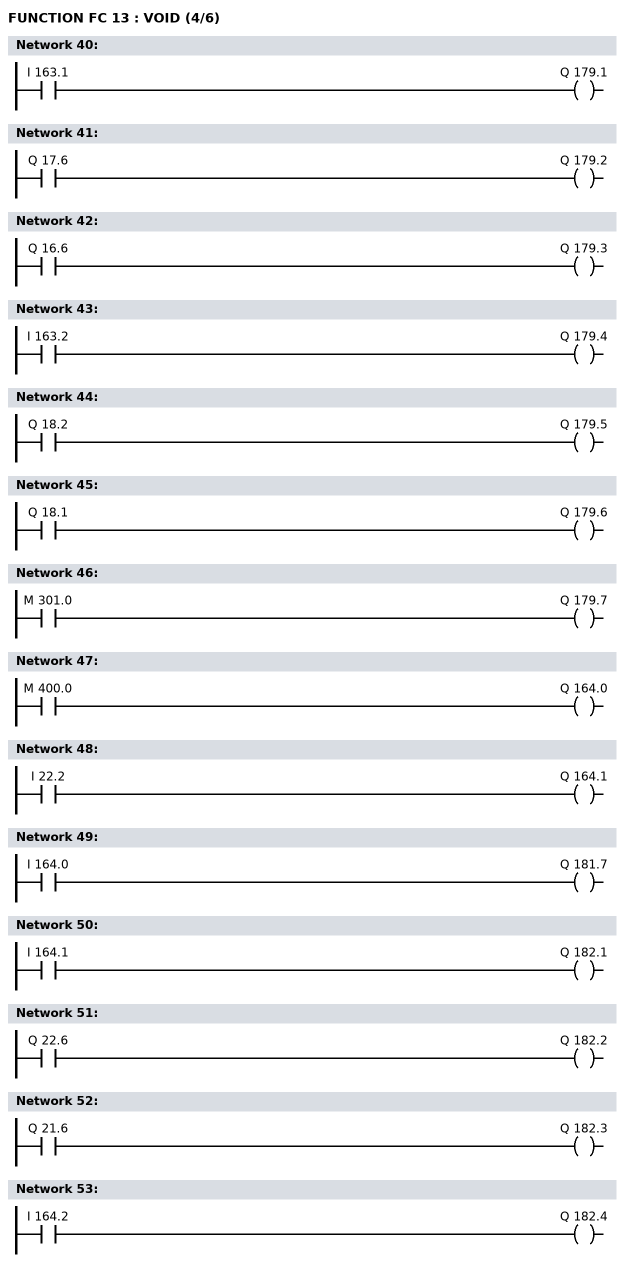

      A     I    163.1;
      =     Q    179.1;
NETWORK
TITLE =

      A     Q     17.6;
      =     Q    179.2;
NETWORK
TITLE =

      A     Q     16.6;
      =     Q    179.3;
NETWORK
TITLE =

      A     I    163.2;
      =     Q    179.4;
NETWORK
TITLE =

      A     Q     18.2;
      =     Q    179.5;
NETWORK
TITLE =

      A     Q     18.1;
      =     Q    179.6;
NETWORK
TITLE =

      A     M    301.0;
      =     Q    179.7;
NETWORK
TITLE =

      A     M    400.0;
      =     Q    164.0;
NETWORK
TITLE =

      A     I     22.2;
      =     Q    164.1;
NETWORK
TITLE =

      A     I    164.0;
      =     Q    181.7;
NETWORK
TITLE =

      A     I    164.1;
      =     Q    182.1;
NETWORK
TITLE =

      A     Q     22.6;
      =     Q    182.2;
NETWORK
TITLE =

      A     Q     21.6;
      =     Q    182.3;
NETWORK
TITLE =

      A     I    164.2;
      =     Q    182.4;
NETWORK
TITLE =
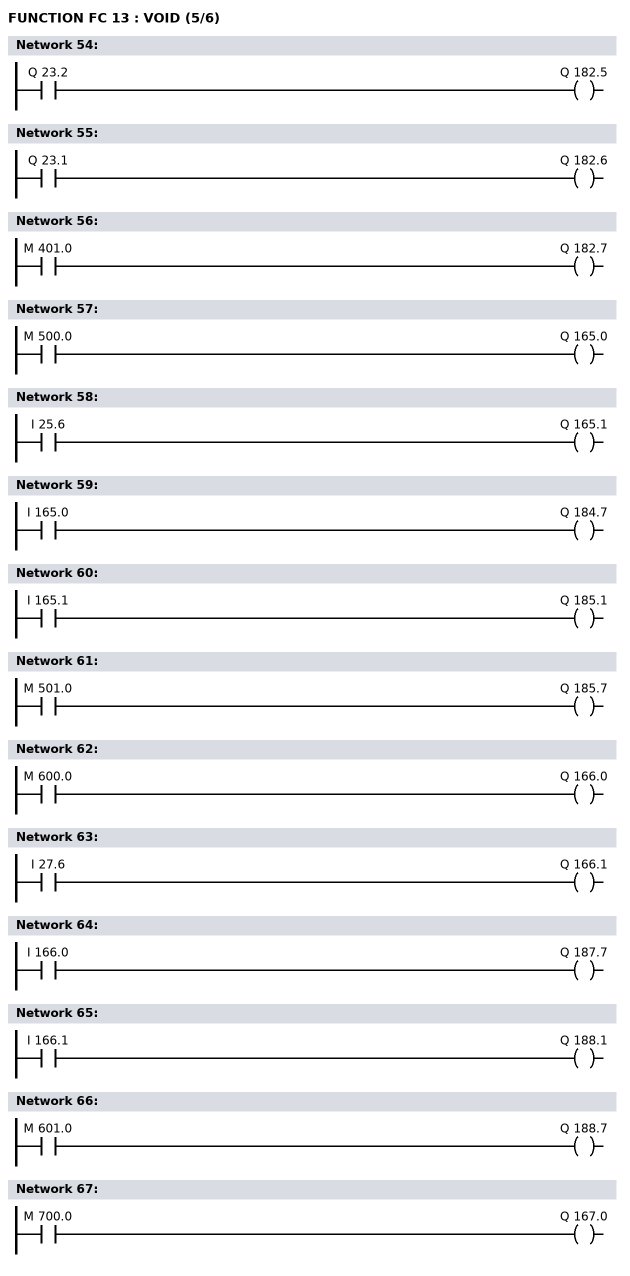

      A     Q     23.2;
      =     Q    182.5;
NETWORK
TITLE =

      A     Q     23.1;
      =     Q    182.6;
NETWORK
TITLE =

      A     M    401.0;
      =     Q    182.7;
NETWORK
TITLE =

      A     M    500.0;
      =     Q    165.0;
NETWORK
TITLE =

      A     I     25.6;
      =     Q    165.1;
NETWORK
TITLE =

      A     I    165.0;
      =     Q    184.7;
NETWORK
TITLE =

      A     I    165.1;
      =     Q    185.1;
NETWORK
TITLE =

      A     M    501.0;
      =     Q    185.7;
NETWORK
TITLE =

      A     M    600.0;
      =     Q    166.0;
NETWORK
TITLE =

      A     I     27.6;
      =     Q    166.1;
NETWORK
TITLE =

      A     I    166.0;
      =     Q    187.7;
NETWORK
TITLE =

      A     I    166.1;
      =     Q    188.1;
NETWORK
TITLE =

      A     M    601.0;
      =     Q    188.7;
NETWORK
TITLE =

      A     M    700.0;
      =     Q    167.0;
NETWORK
TITLE =
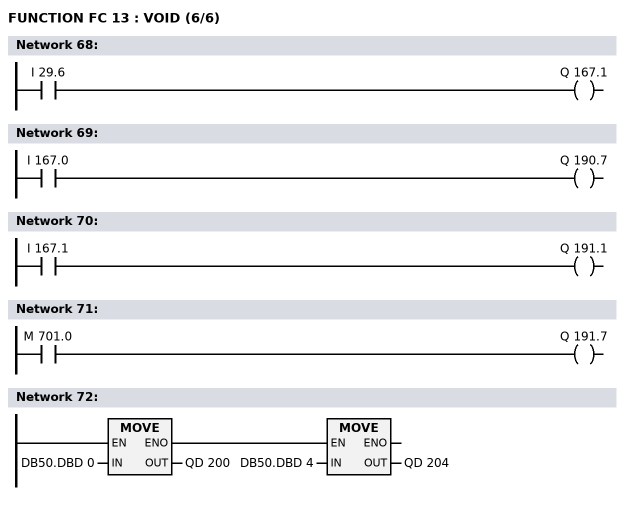

      A     I     29.6;
      =     Q    167.1;
NETWORK
TITLE =

      A     I    167.0;
      =     Q    190.7;
NETWORK
TITLE =

      A     I    167.1;
      =     Q    191.1;
NETWORK
TITLE =

      A     M    701.0;
      =     Q    191.7;
NETWORK
TITLE =

      A(    ;
      L     DB50.DBD    0;
      T     QD   200;
      SET   ;
      SAVE  ;
      CLR   ;
      A     BR;
      )     ;
      JNB   M001;
      L     DB50.DBD    4;
      T     QD   204;
M001: NOP   0;
END_FUNCTION

FUNCTION FC 100 : VOID
VERSION : 0.1

BEGIN
NETWORK
TITLE =
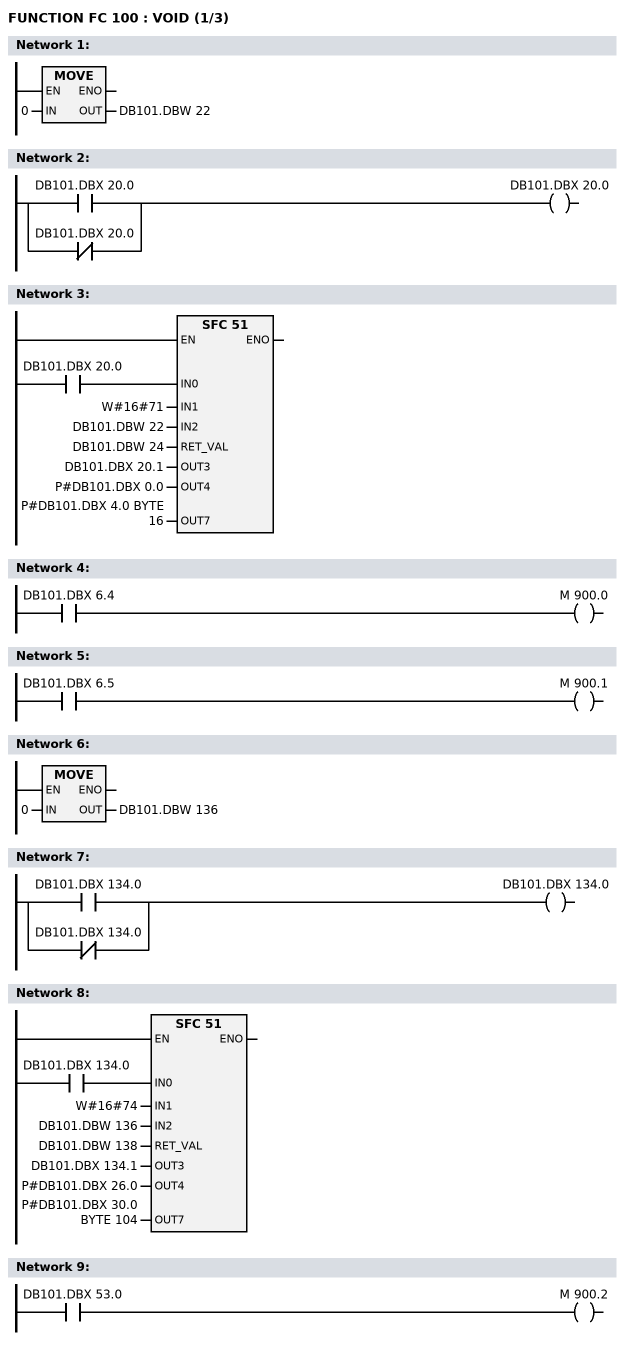

      L     0;
      T     DB101.DBW   22;
      NOP   0;
NETWORK
TITLE =

      O     DB101.DBX   20.0;
      ON    DB101.DBX   20.0;
      =     DB101.DBX   20.0;
NETWORK
TITLE =

      A     DB101.DBX   20.0;
      =     L      0.0;
      BLD   103;
      CALL SFC   51 (
           IN0                      := L      0.0,
           IN1                      := W#16#71,
           IN2                      := DB101.DBW   22,
           RET_VAL                  := DB101.DBW   24,
           OUT3                     := DB101.DBX   20.1,
           OUT4                     := P#DB101.DBX 0.0,
           OUT7                     := P#DB101.DBX 4.0 BYTE 16);
      NOP   0;
NETWORK
TITLE =

      A     DB101.DBX    6.4;
      =     M    900.0;
NETWORK
TITLE =

      A     DB101.DBX    6.5;
      =     M    900.1;
NETWORK
TITLE =

      L     0;
      T     DB101.DBW  136;
      NOP   0;
NETWORK
TITLE =

      O     DB101.DBX  134.0;
      ON    DB101.DBX  134.0;
      =     DB101.DBX  134.0;
NETWORK
TITLE =

      A     DB101.DBX  134.0;
      =     L      0.0;
      BLD   103;
      CALL SFC   51 (
           IN0                      := L      0.0,
           IN1                      := W#16#74,
           IN2                      := DB101.DBW  136,
           RET_VAL                  := DB101.DBW  138,
           OUT3                     := DB101.DBX  134.1,
           OUT4                     := P#DB101.DBX 26.0,
           OUT7                     := P#DB101.DBX 30.0 BYTE 104);
      NOP   0;
NETWORK
TITLE =

      A     DB101.DBX   53.0;
      =     M    900.2;
NETWORK
TITLE =
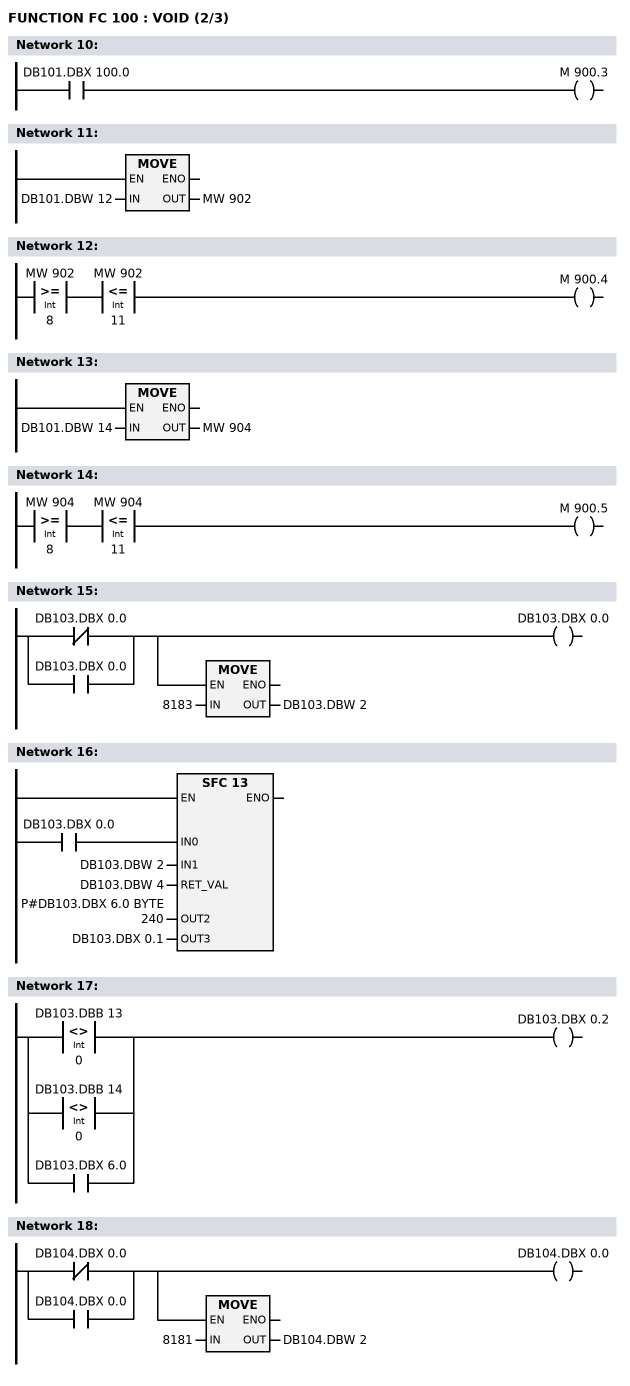

      A     DB101.DBX  100.0;
      =     M    900.3;
NETWORK
TITLE =

      L     DB101.DBW   12;
      T     MW   902;
      NOP   0;
NETWORK
TITLE =

      A(    ;
      L     MW   902;
      L     8;
      >=I   ;
      )     ;
      A(    ;
      L     MW   902;
      L     11;
      <=I   ;
      )     ;
      =     M    900.4;
NETWORK
TITLE =

      L     DB101.DBW   14;
      T     MW   904;
      NOP   0;
NETWORK
TITLE =

      A(    ;
      L     MW   904;
      L     8;
      >=I   ;
      )     ;
      A(    ;
      L     MW   904;
      L     11;
      <=I   ;
      )     ;
      =     M    900.5;
NETWORK
TITLE =

      ON    DB103.DBX    0.0;
      O     DB103.DBX    0.0;
      =     L      0.0;
      A     L      0.0;
      BLD   102;
      =     DB103.DBX    0.0;
      A     L      0.0;
      JNB   M001;
      L     8183;
      T     DB103.DBW    2;
M001: NOP   0;
NETWORK
TITLE =

      A     DB103.DBX    0.0;
      =     L      0.0;
      BLD   103;
      CALL SFC   13 (
           IN0                      := L      0.0,
           IN1                      := DB103.DBW    2,
           RET_VAL                  := DB103.DBW    4,
           OUT2                     := P#DB103.DBX 6.0 BYTE 240,
           OUT3                     := DB103.DBX    0.1);
      NOP   0;
NETWORK
TITLE =

      O(    ;
      L     DB103.DBB   13;
      L     0;
      <>I   ;
      )     ;
      O(    ;
      L     DB103.DBB   14;
      L     0;
      <>I   ;
      )     ;
      O     DB103.DBX    6.0;
      =     DB103.DBX    0.2;
NETWORK
TITLE =

      ON    DB104.DBX    0.0;
      O     DB104.DBX    0.0;
      =     L      0.0;
      A     L      0.0;
      BLD   102;
      =     DB104.DBX    0.0;
      A     L      0.0;
      JNB   M002;
      L     8181;
      T     DB104.DBW    2;
M002: NOP   0;
NETWORK
TITLE =
